(* IEC 61131-3 sources: volt/packages/volt-lsp-iec/test-corpus/lenze-mid/Device/Plc Logic/Application/A70_MachineModuleSources/MM_MachineControl/02_subMain, 11 files *)

(* ---- SidecorrectionCalculation.pou ---- *)
FUNCTION SidecorrectionCalculation
VAR_INPUT
	iAnalogInputValue						: INT;
	iSetpoint								: INT;
	iCorrectionScale						: REAL;
	iLightValue								: INT;
	iDarkValue								: INT;
	iNoWrapperOffsetPercentage01Perc		: INT; //test5

END_VAR
VAR_OUTPUT
	oIntPercentage							: INT;
	oRealPercentage							: REAL;
	oCorrectionValue						: REAL;
	oDeviationNoWrapper						: REAL;
END_VAR
VAR

	tRealMeasuredValue						: REAL;
	tRealPercentage							: REAL;
	tRealSetpoint							: REAL;
	tWhiteValue								: DINT;
	tBrownValue								: DINT;
	tWidthLight_Dark						: DINT;
	tRealWidthLight_Dark					: REAL;
	tMeasuredWithOffset						: REAL;
	tRealBrownValue							: REAL;
	tRealNoWrapperOffsetPercentage			: REAL;

END_VAR

%LANGUAGE ST
//Read out values for light and dark
tWhiteValue:=MOVE(iLightValue);
tBrownValue:=MOVE(iDarkValue);

//Calculate difference between light and dark value (light will be higher than dark)
tRealWidthLight_Dark:=TO_REAL(tWhiteValue-tBrownValue);
tRealBrownValue:=TO_REAL(tBrownValue);

//Measured value compensated with offset
tRealMeasuredValue:=TO_REAL(iAnalogInputValue);
tMeasuredWithOffset:=tRealMeasuredValue-tRealBrownValue;

//Calculation of the percentage
//"Measured value"/ Bandwidth
IF tRealWidthLight_Dark=0 THEN
	tRealWidthLight_Dark:=10;

END_IF
oRealPercentage:=(tMeasuredWithOffset/tRealWidthLight_Dark)*100;
oIntPercentage:=TO_INT(oRealPercentage);

//Calculation of the fault
//(act - set) * "correction scale"
tRealSetpoint:=TO_REAL(iSetpoint);
oCorrectionValue:=(oRealPercentage-tRealSetpoint)*iCorrectionScale;

//No wrapper detection
tRealNoWrapperOffsetPercentage:=TO_REAL(iNoWrapperOffsetPercentage01Perc);
oDeviationNoWrapper:=TO_INT(tRealNoWrapperOffsetPercentage*(tRealWidthLight_Dark/1000));

END_FUNCTION

(* ---- SpeedCalculationTrayfiller.pou ---- *)
FUNCTION SpeedCalculationTrayfiller
VAR_INPUT
END_VAR
VAR
	tInt: INT;
	tBool: BOOL;
END_VAR

%LANGUAGE LD
%NETWORK "NETWORK 1: Write setpoint speed in DB"
// The speed of the trayfiller has to be higher then the speed of the dryer. In this way there is always an empty space at the startpostition of the trayfiller.
MOVE(EN := ADD(EN := RAIL(), Mach1_Data.Drives.FeedForwardADS.Control.AutoSpeed, 30, OUT => tInt), tInt, OUT => Mach1_Data.Drives.FeedForwardATF.Control.AutoSpeed);
%NETWORK "NETWORK 2: Activation + Runtime guard feed forward dryer/trayfiller"
// Runtime calculation:
// 1 cycle = 60s/rpm
// speed = in 0.1 rpm -> 60s = 600 1/10s
//
// -> 1 cycle = 600/speed01
// DINT cannot calculate this 600/1000 = 0.1 -> DINT=0
// First multiply by 1000 (s -> ms)
// 1cycle = (600*1000)/speed1
// To give a little margin: add 500ms
ASSIGN(RuntimeGuard_V5_1_100(AlarmDB := Mach1_Alarms, iForward := Mach1_AuxData.TrayfillerActive AND Mach1_MIDS.IDB_TrayFiller.oFeedForwardMotor AND Mach1.Genflags.DelayAfterSTO AND (Mach1_AuxData.AllDrivesHomed OR INVERT(Mach1_AuxData.TrayfillerActive)), iReverse := LST_General.AlwaysOff, iActivateGuard := GE(EN := Mach1.Genflags.DelayAfterSTO AND Mach1_Data.Drives.FeedForwardATF.Control.StartAuto AND INVERT(LST_InputsOutputs.I133_3_PROX_zero_position_transport_ATF), Mach1_Data.Drives.FeedForwardATF.Control.AutoSpeed, 10).OUT, iMaxRuntime := T#10S, iReset := Mach1.GenFlags.StartFlag, iAlm := Mach1_Alarms.Alm051, ioAction := Mach1.GenFlags.MinorAlarm, ioAccRuntime := Mach1_AuxData.IEC_TIMERS.RuntimeGuardFeedforwardTrayfiller, oForwardGuarded => Mach1_Data.Drives.FeedForwardATF.Control.StartAuto), Q_SET => Mach1.GenFlags.StopDriveDirect);

END_FUNCTION

(* ---- Servo_LimitJog.pou ---- *)
FUNCTION_BLOCK Servo_LimitJog
VAR_INPUT
	iServoStatus 	: sUDT_ServoComm_Drive_Status;
	iServoControl 		: sUDT_ServoComm_Drive_Control;
END_VAR
VAR_OUTPUT
	oServoControl 		: sUDT_ServoComm_Drive_Control;
END_VAR
VAR
END_VAR
VAR_IN_OUT
	ioUDT_ServoDrive			: UDT_ServoDrive;
	ioUDT_JogLimitFree			: UDT_ServoJogLimitFree;
END_VAR

%LANGUAGE LD
%NETWORK "NETWORK 3 (p1): Check for limit switch"
ASSIGN(iServoStatus.Spare1, Q => ioUDT_JogLimitFree.Status.Limit_Left_OK);
%NETWORK "NETWORK 3 (p2): Check for limit switch"
ASSIGN(iServoStatus.Spare2, Q => ioUDT_JogLimitFree.Status.Limit_Right_OK);
%NETWORK "COPY previous control word to current controlword"
EXECUTE(EN := RAIL(), 'oServoControl:=iServoControl;');
%NETWORK "NETWORK 4 (p1): ControlToFreeLimitSwitches"
ASSIGN(ioUDT_JogLimitFree.Status.Limit_Left_OK AND ioUDT_JogLimitFree.Control.Jog_LimitToLeft, Q => oServoControl.Spare1);
%NETWORK "NETWORK 4 (p2): ControlToFreeLimitSwitches"
ASSIGN(ioUDT_JogLimitFree.Status.Limit_Right_OK AND ioUDT_JogLimitFree.Control.Jog_LimitToRight, Q => oServoControl.Spare2);

END_FUNCTION_BLOCK

(* ---- WSM.pou ---- *)
FUNCTION_BLOCK WSM
VAR_INPUT
	EN: BOOL;
	iGenflags : UDT_GeneralFlags;
	iInit: BOOL;
	iTest_Prod: BOOL;
	iCleaning: BOOL;
	iBunchPresent: BOOL;
	iWrapperPresentForLeafCarrier: BOOL;
	iPhotocellWrapper: BOOL;
	iWaterLevelSensor: BOOL;
	iTakeOverCycle: BOOL;
	iTimeOutSupplyWrapper: TIME;
	iSprayTime: TIME;
	iDelayContSpraying: TIME;
	iScreenForOperatorSettingsActivated: BOOL;
	iManualSprayCycleReset: BOOL;
	iManualSprayCycleStart: BOOL;
	iManualSprayCycleStop: BOOL;
	iMaxNumberOfSprayPulses: INT;

END_VAR
VAR_OUTPUT
	ENO: BOOL;
	oVentilationMotor: BOOL;
	oPositionMotor: BOOL;
	oWindingMotor: BOOL;
	oSprayingValve: BOOL;
	oWaterLevelValve: BOOL;
	oFaultWaitingForWrapper: BOOL;
	oFaultNoWrapper: BOOL;
	oFaultPhotocellWrapper : BOOL;
END_VAR
VAR
	stOSN_TakeOverCycle: F_TRIG;
	TMR_TimeOutSupply: TON;
	TMR_TimeOutPhotocell: TON;
	stRePositionMotor: R_TRIG;
	stSprayCycleActive: BOOL;
	TMR_DelayContinuousSpraying: TON;
	TMR_SprayTime: TON;
	stManualSprayCycleStarted: BOOL;

	TMR_ManualSprayCycleIdle: TON;

END_VAR

VAR_IN_OUT
	ioEnableSpraying: BOOL;
	ioManualSprayCycleActualCount: INT;
	ioManualStartSupply: BOOL;
END_VAR
VAR RETAIN PERSISTENT
	stRestposition: BOOL;
	stSupplyWrapper: BOOL;
	stWrapperPresent: BOOL;
	stNoWrapper: BOOL;
	stPhotocellWrapperFault: BOOL;
	stFeedForward: BOOL;
END_VAR
%LANGUAGE LD
%NETWORK "DONE Network 2: State: Initialise"
VAR w1 : ANY; END_VAR
w1 := iInit OR INVERT(iTest_Prod) OR iCleaning OR ioManualStartSupply;
ASSIGN(w1, Q_SET => stRestposition);
ASSIGN(w1, Q_RESET => stSupplyWrapper, Q_RESET => stWrapperPresent, Q_RESET => stNoWrapper, Q_RESET => stPhotocellWrapperFault);
%NETWORK "DONE Network 3: State: Restposition"
ASSIGN(stOSN_TakeOverCycle(CLK := iTakeOverCycle) AND stWrapperPresent, Q_SET => stRestposition, Q_RESET => stWrapperPresent);
%NETWORK "DONE Network 4: State: Supply wrapper"
ASSIGN(stRestposition AND (iTest_Prod AND INVERT(iCleaning) AND iBunchPresent AND INVERT(iTakeOverCycle) AND (iGenFlags.RunMan OR iGenFlags.RunAuto) OR ioManualStartSupply) OR stNoWrapper AND iGenFlags.StartFlag OR stPhotocellWrapperFault AND iGenFlags.StartFlag, Q_SET => stSupplyWrapper, Q_RESET => stRestposition, Q_RESET => stNoWrapper, Q_RESET => stPhotocellWrapperFault, Q_RESET => ioManualStartSupply);
%NETWORK "DONE Network 5: State: Wrapper Present"
VAR w2 : ANY; END_VAR
w2 := iWrapperPresentForLeafCarrier AND stSupplyWrapper;
ASSIGN(w2, Q_SET => stWrapperPresent);
ADD(EN := w2, 1, HMI_Var.Mach1.PRDWrapCurrentCntr, OUT => HMI_Var.Mach1.PRDWrapCurrentCntr);
ADD(EN := w2, 1, HMI_Var.Mach1.PRDWrapDayCounter, OUT => HMI_Var.Mach1.PRDWrapDayCounter);
ASSIGN(w2, Q_RESET => stSupplyWrapper);
%NETWORK "DONE Network 6: State: No Wrapper"
ASSIGN(TMR_TimeOutSupply(IN := stSupplyWrapper AND stFeedForward, PT := iTimeOutSupplyWrapper), Q_SET => stNoWrapper, Q_RESET => stSupplyWrapper);
%NETWORK "DONE Network 7: State: Photocell wrapper fault"
ASSIGN(TMR_TimeOutPhotocell(IN := stSupplyWrapper AND stFeedForward AND iPhotocellWrapper, PT := T#10S), Q_SET => stPhotocellWrapperFault, Q_RESET => stSupplyWrapper);
%NETWORK "DONE Network 8: Faults"
VAR w3 : ANY; END_VAR
w3 := True;
ASSIGN(w3 AND stSupplyWrapper AND iTakeOverCycle, Q => oFaultWaitingForWrapper);
ASSIGN(w3 AND stNoWrapper, Q => oFaultNoWrapper);
ASSIGN(w3 AND stPhotocellWrapperFault, Q => oFaultPhotocellWrapper);
%NETWORK "DONE Network 9: Ventilation motor"
ASSIGN(iGenFlags.EnableAuxDrive AND iTest_Prod AND INVERT(iCleaning), Q => oVentilationMotor);
%NETWORK "DONE Network 10:"
VAR w4 : ANY; END_VAR
w4 := iGenFlags.EnableAuxDrive AND stSupplyWrapper AND INVERT(iGenFlags.StopFlag);
ASSIGN(w4, Q => stFeedForward);
ASSIGN(w4, Q => oPositionMotor);
%NETWORK "DONE Network 11: Winding motor"
ASSIGN(iGenFlags.EnableAuxDrive AND INVERT(iGenFlags.StopFlag) AND iTest_Prod AND INVERT(iCleaning), Q => oWindingMotor);
%NETWORK "DONE Network 12: Start spray cycle"
VAR w5 : ANY; END_VAR
w5 := stFeedForward;
ASSIGN(stRePositionMotor(CLK := w5), Q_SET => stSprayCycleActive);
ASSIGN(TMR_DelayContinuousSpraying(IN := w5, PT := iDelayContSpraying), Q_SET => stSprayCycleActive);
%NETWORK "DONE Network 13: Timing spray cycle"
ASSIGN(TMR_SprayTime(IN := stSprayCycleActive, PT := iSprayTime) AND INVERT(TMR_DelayContinuousSpraying.Q), Q_RESET => stSprayCycleActive);
%NETWORK "DONE Network 14: Spraying valve"
ASSIGN(ioEnableSpraying AND stSprayCycleActive, Q => oSprayingValve);
%NETWORK "DONE Network 15: Automatic trigger of water"
ASSIGN(FALSE AND iGenFlags.EnablePneumEStop AND iWrapperPresentForLeafCarrier AND iTest_Prod AND INVERT(iCleaning), Q_SET => ioEnableSpraying);
%NETWORK "DONE Network 16: Water level control"
ASSIGN(ioEnableSpraying AND iWaterLevelSensor, Q => oWaterLevelValve);
%NETWORK "DONE Network 17: Manual spray cycle"
VAR w6 : ANY; END_VAR
w6 := iScreenForOperatorSettingsActivated;
MOVE(EN := w6 AND iManualSprayCycleReset, 0, OUT => ioManualSprayCycleActualCount);
ASSIGN(LT(EN := w6 AND iGenFlags.EnablePneumEStop AND (iManualSprayCycleStart OR stManualSprayCycleStarted) AND INVERT(iManualSprayCycleStop) AND INVERT(iManualSprayCycleReset), ioManualSprayCycleActualCount, iMaxNumberOfSprayPulses).OUT, Q => stManualSprayCycleStarted);
ASSIGN(ADD(EN := TMR_ManualSprayCycleIdle(IN := w6 AND stManualSprayCycleStarted AND INVERT(stSprayCycleActive), PT := T#300MS), ioManualSprayCycleActualCount, 1, OUT => ioManualSprayCycleActualCount), Q_SET => stSprayCycleActive);
%NETWORK "DONE Network 18: SAVE RLO"
ASSIGN(EN, Q => ENO);

END_FUNCTION_BLOCK

(* ---- AHWF.pou ---- *)
PROGRAM AHWF
VAR
	tFaultWaitingForWrapper : BOOL;
	tFaultNoWrapper: BOOL;
	tFaultPhotocellWrapper: BOOL;
	tStartFastWinding: BOOL;
	tSupplyWrapper: BOOL;
	tSprayingValve: BOOL;
	ttest: BOOL;
	R_TrigStartPos: R_TRIG;
END_VAR

VAR
	IDB_WSM: WSM;
END_VAR
%LANGUAGE LD
%NETWORK "Network 1: Detection of wrapper (set and reset)"
VAR w1 : ANY; END_VAR
w1 := True;
ASSIGN(w1 AND LST_InputsOutputs.I101_0_Wrapper_present, Q_SET => Mach1_AuxData.MemWrapperPassedUnderTheSensor);
ASSIGN(w1 AND INVERT(LST_InputsOutputs.I101_0_Wrapper_present) AND Mach1_AuxData.MemWrapperPassedUnderTheSensor, Q_SET => Mach1_AuxData.MemWrapperPresentForLeafCarrier, Q_SET => Mach1_AuxData.MemWrapperDetected_ResetLimitedSpeed);
ASSIGN(fc_CamC_CP_UDT(iEN := MOVE(EN := w1, Mach1_Data.CamControls.TakeOverCycle_C.Stop, OUT => Mach1_AuxData.CamControls.TakeOverCycleStopPulse_CP.Start), iMachinePosition := HMI_Var.Mach1.Position, iResetFlag := Mach1.GenFlags.Rotflag, ioPulse := Mach1_AuxData.CamControls.TakeOverCycleStopPulse_CP), Q_RESET => Mach1_AuxData.MemWrapperPresentForLeafCarrier, Q_RESET => Mach1_AuxData.MemWrapperPassedUnderTheSensor);
%NETWORK
ASSIGN(R_TrigStartPos(CLK := HMI_Var.HMI_AHWF_StartPos), Q_RESET => Mach1_AuxData.MemWrapperPresentForLeafCarrier, Q_RESET => Mach1_AuxData.MemWrapperPassedUnderTheSensor);
%NETWORK "Network 2: FB for DTA"
ASSIGN(IDB_WSM(EN := RAIL(), iGenflags := Mach1.GenFlags, iInit := LST_General.FirstCycle, iTest_Prod := HMI_Var.Test_Prod, iCleaning := HMI_Var.Btn_Cleaning, iBunchPresent := Mach1_AuxData.ShiftRegister.SR_bunch_present_position_1_JL, iWrapperPresentForLeafCarrier := Mach1_AuxData.MemWrapperPresentForLeafCarrier AND INVERT(HMI_Var.HMI_AHWF_fast_winding), iPhotocellWrapper := LST_InputsOutputs.I101_0_Wrapper_present AND INVERT(HMI_Var.HMI_AHWF_fast_winding), iWaterLevelSensor := LST_InputsOutputs.I101_3_Water_level_control, iTakeOverCycle := fc_CamC_CC_UDT(iEnable := True, iMachinePosition := HMI_Var.Mach1.Position, ioCamControl := Mach1_Data.CamControls.TakeOverCycle_C), iTimeOutSupplyWrapper := OPERAND('fc_dinttotime(Mach1_Data.Timers.TimeOutSupplyWrapper,2)'), iSprayTime := OPERAND('fc_dinttotime(Mach1_Data.Timers.SprayPulseWidth,2)'), iDelayContSpraying := OPERAND('fc_dinttotime(Mach1_Data.Timers.DelayContSpraying,2)'), iScreenForOperatorSettingsActivated := Mach1_AuxData.ScreenForOperatorSettingsActivated, iManualSprayCycleReset := HMI_Var.Mach1.SprayReset, iManualSprayCycleStart := HMI_Var.Mach1.SprayStart, iManualSprayCycleStop := HMI_Var.Mach1.SprayStop, iMaxNumberOfSprayPulses := Mach1_Data.Settings.Ints.MaxNumberOfSprayPulses, ioEnableSpraying := HMI_Var.Btn_Spraying, ioManualSprayCycleActualCount := Mach1_Data.Settings.Ints.ActualNumberOfSprayPulses, ioManualStartSupply := HMI_Var.HMI_AHWF_StartPos, oPositionMotor => tSupplyWrapper, oSprayingValve => tSprayingValve, oWaterLevelValve => LST_InputsOutputs.Q101_1_PNV_Waterlevel_control, oFaultWaitingForWrapper => tFaultWaitingForWrapper, oFaultNoWrapper => tFaultNoWrapper, oFaultPhotocellWrapper => tFaultPhotocellWrapper) AND Mach1.GenFlags.EnablePneumPressurised AND Mach1_Safety.Status.AllDoorsActuallyClosed AND tSprayingValve AND INVERT(Mach1_Alarms.Alm011), Q => PneumValveTerminalSMC.Pos1B);
%NETWORK "Network 3: Wrapper faults"
ASSIGN(Alarms_V5_1_100(AlarmDB := Mach1_Alarms, iCond := Mach1.GenFlags.DelayAfterEmergStop AND HMI_Var.Test_Prod AND INVERT(HMI_Var.Btn_Cleaning) AND tFaultWaitingForWrapper AND Mach1_AuxData.AllDrivesHomed, iReset := True, iAlm := Mach1_Alarms.Alm076, ioAction := Mach1.GenFlags.Warning) OR Alarms_V5_1_100(AlarmDB := Mach1_Alarms, iCond := Mach1.GenFlags.DelayAfterEmergStop AND HMI_Var.Test_Prod AND INVERT(HMI_Var.Btn_Cleaning) AND tFaultNoWrapper AND Mach1_AuxData.AllDrivesHomed, iReset := Mach1.GenFlags.StartFlag, iAlm := Mach1_Alarms.Alm043, ioAction := Mach1.GenFlags.MinorAlarm) OR Alarms_V5_1_100(AlarmDB := Mach1_Alarms, iCond := Mach1.GenFlags.DelayAfterEmergStop AND HMI_Var.Test_Prod AND INVERT(HMI_Var.Btn_Cleaning) AND INVERT(Mach1_Alarms.Alm045) AND tFaultPhotocellWrapper AND Mach1_AuxData.AllDrivesHomed, iReset := Mach1.GenFlags.StartFlag, iAlm := Mach1_Alarms.Alm045, ioAction := Mach1.GenFlags.MinorAlarm), Q_SET => Mach1.GenFlags.StopDriveDirect);
%NETWORK
%NETWORK "TODO Network 4: "
VAR w2 : ANY; w3 : ANY; w4 : ANY; END_VAR
w2 := True;
w3 := w2 AND True;
MOVE(EN := MOVE(EN := MOVE(EN := MOVE(EN := w3 AND TRUE, 175, OUT => Data_Exchange_Motion.FeedForwardWrapper.Control.VelUnit), 2000, OUT => Data_Exchange_Motion.FeedForwardWrapper.Control.DecUnit), 750, OUT => Data_Exchange_Motion.FeedForwardWrapper.Control.AccUnit), 100, OUT => Data_Exchange_Motion.FeedForwardWrapper.Control.TorqueLimit);
w4 := w3 AND HMI_Var.HMI_AHWF_fast_winding;
ASSIGN(Mach1_AuxData.IEC_TIMERS.TON_StartFastWinding(IN := w4, PT := T#200MS), Q => tStartFastWinding);
MOVE(EN := w4, 500, OUT => Data_Exchange_Motion.FeedForwardWrapper.Control.VelUnit);
MOVE(EN := w2, OPERAND('DINT_TO_LREAL(Mach1_Data.Settings.Dints.WrapperStopPosition)/10'), OUT => Data_Exchange_Motion.FeedForwardWrapper.Control.PosUnit);
ASSIGN(w2 AND INVERT(HMI_Var.HMI_AHWF_positioningType) AND INVERT(Mach1_Alarms.Alm056) AND mach1.Genflags.EnableAuxDrive AND (tSupplyWrapper OR tStartFastWinding OR Data_Exchange_Motion.FeedForwardWrapper.Control.StartTouchprobePos AND INVERT(Data_Exchange_Motion.FeedForwardWrapper.Status.InPosition)), Q => Data_Exchange_Motion.FeedForwardWrapper.Control.StartTouchprobePos);
ASSIGN(Mach1_AuxData.Edge.OSP_StopFlag(CLK := w2 AND (INVERT(Mach1_MIDS.FB_Mach1.iStop1) OR INVERT(Mach1_MIDS.FB_Mach1.iStop2) OR INVERT(Mach1_MIDS.FB_Mach1.iStop3) OR INVERT(Mach1_Safety.Status.AllDoorsActuallyClosed) OR LST_InputsOutputs.I101_0_Wrapper_present)), Q_RESET => HMI_Var.HMI_AHWF_fast_winding);
%NETWORK "Network 5: Side correction"
SideCorrection(EN := RAIL());
%NETWORK "Network 6: DTA-alarm: side limit reached"
ASSIGN(Alarms_V5_1_100(AlarmDB := Mach1_Alarms, iCond := Mach1_AuxData.Edge.OSP_LimitDTA_Reached(CLK := Mach1_AuxData.MIDS_Active AND Mach1.GenFlags.DelayAfterEmergStop AND (INVERT(Mach1_Data.Drives.SideCorrection_FreeLimit.Status.Limit_Left_OK) OR INVERT(Mach1_Data.Drives.SideCorrection_FreeLimit.Status.Limit_Right_OK))) AND Mach1_AuxData.AllDrivesHomed, iReset := Mach1.GenFlags.StartFlag, iAlm := Mach1_Alarms.Alm057, ioAction := Mach1.GenFlags.MinorAlarm) OR LST_General.AlwaysOff AND Alarms_V5_1_100(AlarmDB := Mach1_Alarms, iCond := Mach1_AuxData.MIDS_Active AND Mach1.GenFlags.DelayAfterEmergStop AND (INVERT(Mach1_Data.Drives.SideCorrection_FreeLimit.Status.Limit_Left_OK) OR INVERT(Mach1_Data.Drives.SideCorrection_FreeLimit.Status.Limit_Right_OK)) AND Mach1_AuxData.AllDrivesHomed, iReset := Mach1.GenFlags.StartFlag, iAlm := Mach1_Alarms.Alm074, ioAction := Mach1.GenFlags.Warning), Q_SET => Mach1.GenFlags.StopDriveDirect);
%NETWORK "Network 7: Alarm: Water receptacle full"
ASSIGN(Alarms_V5_1_100(AlarmDB := Mach1_Alarms, iCond := Mach1_AuxData.IEC_TIMERS.WaterReceptacleFull(IN := Mach1_AuxData.MIDS_Active AND LST_InputsOutputs.I101_3_Water_level_control AND INVERT(Mach1_Alarms.Alm055), PT := T#5M) AND HMI_Var.Test_Prod AND HMI_Var.Btn_Spraying AND Mach1_AuxData.AllDrivesHomed, iReset := Mach1.GenFlags.StartFlag, iAlm := Mach1_Alarms.Alm055, ioAction := Mach1.GenFlags.MinorAlarm), Q_SET => Mach1.GenFlags.StopDriveDirect);

END_PROGRAM

(* ---- fc_CheckRegister.pou ---- *)
PROGRAM fc_CheckRegister
VAR
END_VAR

%LANGUAGE LD
%NETWORK "NETWORK 1: Shift CheckRegister"
fc_ShiftRegister(ioPositie := db_CheckRegister.Positie);
%NETWORK "NETWORK 2: Check for error in dryer"
fc_CheckNumberOfErrorsRegister(iPositie := db_CheckRegister.Positie, iPositionToCheck := CTE.posCigarPresentOutfeed, iAmountOfErrors := Mach1_Data.Counters.MaxRepetitionNoCigarsDryer.SetValue, oError => db_CheckRegister.CheckRegisterError);

END_PROGRAM

(* ---- fc_Visualisation_HMI.pou ---- *)
PROGRAM fc_Visualisation_HMI
VAR_INPUT
END_VAR
VAR
	tbool: BOOL;
END_VAR

%LANGUAGE LD
%NETWORK "NETWORK 5: (P1) Visualisation - emergency stop"
Alarms_V5_1_100(AlarmDB := Mach1_Alarms, iCond := Mach1_AuxData.MIDS_Active AND INVERT(Mach1_Safety.Status.Emergency_button01), iReset := True, iAlm := Mach1_Alarms.Alm080, ioAction := Mach1.GenFlags.warning);
%NETWORK "NETWORK 5: (P2) Visualisation - emergency stop"
Alarms_V5_1_100(AlarmDB := Mach1_Alarms, iCond := Mach1_AuxData.MIDS_Active AND INVERT(Mach1_Safety.Status.Emergency_button02), iReset := True, iAlm := Mach1_Alarms.Alm081, ioAction := Mach1.GenFlags.warning);
%NETWORK "NETWORK 5: (P3) Visualisation - emergency stop"
Alarms_V5_1_100(AlarmDB := Mach1_Alarms, iCond := Mach1_AuxData.MIDS_Active AND INVERT(Mach1_Safety.Status.Emergency_button04), iReset := True, iAlm := Mach1_Alarms.Alm082, ioAction := Mach1.GenFlags.warning);
%NETWORK "DONE NETWORK 5 (p2): Visualisation - doors"
ASSIGN(Alarms_V5_1_100(AlarmDB := Mach1_Alarms, iCond := Mach1_AuxData.MIDS_Active AND Mach1.Genflags.DelayAfterEmergStop AND INVERT(Mach1_Safety.Status.Door_switch01), iReset := True, iAlm := Mach1_Alarms.Alm083, ioAction := Mach1.GenFlags.warning) OR Alarms_V5_1_100(AlarmDB := Mach1_Alarms, iCond := Mach1_AuxData.MIDS_Active AND Mach1.Genflags.DelayAfterEmergStop AND INVERT(Mach1_Safety.Status.Door_switch02), iReset := True, iAlm := Mach1_Alarms.Alm084, ioAction := Mach1.GenFlags.warning) OR Alarms_V5_1_100(AlarmDB := Mach1_Alarms, iCond := Mach1_AuxData.MIDS_Active AND Mach1.Genflags.DelayAfterEmergStop AND INVERT(Mach1_Safety.Status.Door_switch03), iReset := True, iAlm := Mach1_Alarms.Alm085, ioAction := Mach1.GenFlags.warning) OR Alarms_V5_1_100(AlarmDB := Mach1_Alarms, iCond := Mach1_AuxData.MIDS_Active AND Mach1.Genflags.DelayAfterEmergStop AND INVERT(Mach1_Safety.Status.Door_switch04), iReset := True, iAlm := Mach1_Alarms.Alm086, ioAction := Mach1.GenFlags.warning) OR Alarms_V5_1_100(AlarmDB := Mach1_Alarms, iCond := Mach1_AuxData.MIDS_Active AND Mach1.Genflags.DelayAfterEmergStop AND INVERT(Mach1_Safety.Status.Door_switch05), iReset := True, iAlm := Mach1_Alarms.Alm087, ioAction := Mach1.GenFlags.warning), Q => tbool);
%NETWORK
ASSIGN(Alarms_V5_1_100(AlarmDB := Mach1_Alarms, iCond := Mach1_AuxData.MIDS_Active AND Mach1.Genflags.DelayAfterEmergStop AND INVERT(Mach1_Safety.Status.Door_switch06), iReset := True, iAlm := Mach1_Alarms.Alm088, ioAction := Mach1.GenFlags.warning) OR Alarms_V5_1_100(AlarmDB := Mach1_Alarms, iCond := Mach1_AuxData.MIDS_Active AND Mach1.Genflags.DelayAfterEmergStop AND INVERT(Mach1_Safety.Status.Door_switch07), iReset := True, iAlm := Mach1_Alarms.Alm089, ioAction := Mach1.GenFlags.warning) OR Alarms_V5_1_100(AlarmDB := Mach1_Alarms, iCond := Mach1_AuxData.MIDS_Active AND Mach1.Genflags.DelayAfterEmergStop AND INVERT(Mach1_Safety.Status.Door_switch08), iReset := True, iAlm := Mach1_Alarms.Alm090, ioAction := Mach1.GenFlags.warning) OR Alarms_V5_1_100(AlarmDB := Mach1_Alarms, iCond := Mach1_AuxData.MIDS_Active AND Mach1.Genflags.DelayAfterEmergStop AND INVERT(Mach1_Safety.Status.Door_switch09), iReset := True, iAlm := Mach1_Alarms.Alm091, ioAction := Mach1.GenFlags.warning) OR Alarms_V5_1_100(AlarmDB := Mach1_Alarms, iCond := Mach1_AuxData.MIDS_Active AND Mach1.Genflags.DelayAfterEmergStop AND INVERT(Mach1_Safety.Status.Door_switch10), iReset := True, iAlm := Mach1_Alarms.Alm092, ioAction := Mach1.GenFlags.warning), Q => tbool);
%NETWORK
ASSIGN(Alarms_V5_1_100(AlarmDB := Mach1_Alarms, iCond := Mach1_AuxData.MIDS_Active AND Mach1.Genflags.DelayAfterEmergStop AND INVERT(Mach1_Safety.Status.Door_switch14), iReset := True, iAlm := Mach1_Alarms.Alm093, ioAction := Mach1.GenFlags.warning) OR Alarms_V5_1_100(AlarmDB := Mach1_Alarms, iCond := Mach1_AuxData.MIDS_Active AND Mach1.Genflags.DelayAfterEmergStop AND INVERT(Mach1_Safety.Status.Door_switch15), iReset := True, iAlm := Mach1_Alarms.Alm094, ioAction := Mach1.GenFlags.warning) OR Alarms_V5_1_100(AlarmDB := Mach1_Alarms, iCond := Mach1_AuxData.MIDS_Active AND Mach1.Genflags.DelayAfterEmergStop AND INVERT(Mach1_Safety.Status.Door_switch16), iReset := True, iAlm := Mach1_Alarms.Alm095, ioAction := Mach1.GenFlags.warning) OR Alarms_V5_1_100(AlarmDB := Mach1_Alarms, iCond := Mach1_AuxData.MIDS_Active AND Mach1.Genflags.DelayAfterEmergStop AND INVERT(Mach1_Safety.Status.Door_switch11), iReset := True, iAlm := Mach1_Alarms.Alm070, ioAction := Mach1.GenFlags.warning) OR Alarms_V5_1_100(AlarmDB := Mach1_Alarms, iCond := Mach1_AuxData.MIDS_Active AND Mach1.Genflags.DelayAfterEmergStop AND INVERT(Mach1_Safety.Status.Door_switch12), iReset := True, iAlm := Mach1_Alarms.Alm071, ioAction := Mach1.GenFlags.warning), Q => tbool);
%NETWORK
Alarms_V5_1_100(AlarmDB := Mach1_Alarms, iCond := Mach1_AuxData.MIDS_Active AND Mach1.Genflags.DelayAfterEmergStop AND INVERT(Mach1_Safety.Status.Door_switch13), iReset := True, iAlm := Mach1_Alarms.Alm072, ioAction := Mach1.GenFlags.warning);
%NETWORK
ASSIGN(Alarms_V5_1_100(AlarmDB := Mach1_Alarms, iCond := Mach1_AuxData.MIDS_Active AND Mach1.Genflags.DelayAfterEmergStop AND LST_InputsOutputs.I100_3_Selector_switch_auto_manual_OP0a, iReset := True, iAlm := Mach1_Alarms.Alm018, ioAction := Mach1.GenFlags.warning) OR Alarms_V5_1_100(AlarmDB := Mach1_Alarms, iCond := Mach1_AuxData.MIDS_Active AND Mach1.Genflags.DelayAfterEmergStop AND LST_InputsOutputs.I132_3_SW_Auto_Man, iReset := True, iAlm := Mach1_Alarms.Alm019, ioAction := Mach1.GenFlags.warning), Q => tbool);
%NETWORK "Reset of alarmlogging"
ASSIGN(Alarms_ResetAlarmLogging(EN := HMI_Var.ResetAlarmLogging, AlarmDB := Mach1_Alarms), Q_RESET => HMI_Var.ResetAlarmLogging);
%NETWORK "Adding product counters$R$L"
ASSIGN(ADD(EN := ADD(EN := ADD(EN := HMI_Var.Mach1.PRDCounterIncr, HMI_Var.Mach1.PRDTotalCounter, 1, OUT => HMI_Var.Mach1.PRDTotalCounter), HMI_Var.Mach1.PRDCigDayCounter, 1, OUT => HMI_Var.Mach1.PRDCigDayCounter), HMI_Var.Mach1.PRDCigCurrentCntr, 1, OUT => HMI_Var.Mach1.PRDCigCurrentCntr), Q_RESET => HMI_Var.Mach1.PRDCounterIncr);
%NETWORK "Reset Day Counter$R$L"
ASSIGN(MOVE(EN := MOVE(EN := HMI_Var.Mach1.PRDDayCounterReset_01, 0, OUT => HMI_Var.Mach1.PRDWrapDayCounter), 0, OUT => HMI_Var.Mach1.PRDCigDayCounter), Q_RESET => HMI_Var.Mach1.PRDDayCounterReset_01);
%NETWORK "Reset Current Counter$R$L"
ASSIGN(MOVE(EN := MOVE(EN := HMI_Var.Mach1.PRDDayCounterReset, 0, OUT => HMI_Var.Mach1.PRDWrapCurrentCntr), 0, OUT => HMI_Var.Mach1.PRDCigCurrentCntr), Q_RESET => HMI_Var.Mach1.PRDDayCounterReset);
%NETWORK
PRG_AlarmsToDWord(EN := TRUE);

END_PROGRAM

(* ---- MainDrive.pou ---- *)
PROGRAM MainDrive
VAR_INPUT
END_VAR
VAR
	tInt: INT;
	tMainDriveRun: BOOL;
	tMainDriveJog: BOOL;
END_VAR

VAR_OUTPUT
	oMainDriveRun: BOOL;
	oMainDriveJog: BOOL;
END_VAR
%LANGUAGE LD
%NETWORK "DONE NETWORK 1: Delay after doors closed"
ASSIGN(Mach1_AuxData.IEC_TIMERS.TON_DelayAfterDoorsClosed(IN := Mach1.GenFlags.DelayAfterEmergStop AND Mach1_Safety.Status.AllDoorsActuallyClosed AND Mach1_Safety.Status.DoorsOK, PT := T#150MS), Q => Mach1_AuxData.DelayAfterDoorsActuallyClosed);
%NETWORK "DONE NETWORK 2: Activating main drive"
VAR w1 : ANY; w2 : ANY; w3 : ANY; w4 : ANY; END_VAR
w1 := TRUE;
MOVE(EN := w1, 0, OUT => tInt);
ASSIGN(w1 AND INVERT(HMI_Var.Test_Prod), Q_RESET => Mach1_AuxData.MemLowerSpeedBecauseOfNoWrapper);
w2 := w1 AND Mach1.GenFlags.EnableMainDrive AND Mach1.GenFlags.ConditionsReadyForOperation AND INVERT(Mach1.GenFlags.StopDriveDirect) AND Mach1_AuxData.AllDrivesInLock;
w3 := w2 AND Mach1.GenFlags.RunAuto;
ASSIGN(w3, Q => tMainDriveRun, Q => oMainDriveRun, Q => Mach1_Safety.Control.RequestAutoSpeed);
MOVE(EN := BRANCH(FEED := w3, INVERT(Mach1_AuxData.MemLowerSpeedBecauseOfNoWrapper), LE(EN := Mach1_AuxData.MemLowerSpeedBecauseOfNoWrapper, Mach1_Data.AUTOSPEED, 40).OUT) AND INVERT(HMI_Var.Btn_Cleaning), Mach1_Data.AUTOSPEED, OUT => tInt);
MOVE(EN := GT(EN := w3 AND Mach1_AuxData.MemLowerSpeedBecauseOfNoWrapper, Mach1_Data.AUTOSPEED, 40).OUT AND INVERT(HMI_Var.Btn_Cleaning), 30, OUT => tInt);
MOVE(EN := w3 AND HMI_Var.Btn_Cleaning, 6, OUT => tInt);
w4 := w2 AND Mach1.GenFlags.RunMan;
ASSIGN(w4, Q => tMainDriveJog, Q => oMainDriveJog, Q => Mach1_Safety.Control.RequestManSpeed);
MOVE(EN := w4, Mach1_Data.MANUALSPEED, OUT => tInt);
RPM_To_DriveSpeed(iEN := w1, iRPM := tInt, oDriveSpeed => Mach1_Data.Drives.MainDrive_VM.Control.DriveMasterSpeed);
%NETWORK "DONE NETWORK 3 : DriveIsRunning flag"
VAR w5 : ANY; END_VAR
w5 := TRUE;
ASSIGN(w5, Q_RESET => Mach1.GenFlags.StopDriveDirect);
ASSIGN(w5 AND (tMainDriveRun OR tMainDriveJog), Q => Mach1.GenFlags.DriveIsRunning);
ASSIGN(Mach1_AuxData.IEC_TIMERS.TOFF_MainDriveAtProductionSpeed(IN := Mach1_AuxData.IEC_TIMERS.TON_MainDriveAtProductionSpeed(IN := w5 AND tMainDriveRun, PT := T#200MS), PT := T#60MS), Q => Mach1.GenFlags.DriveAtSpeed);
%NETWORK "DONE NETWORK 4: Alarm: Main drive blocked"
ASSIGN(Alarms_V5_1_100(AlarmDB := Mach1_Alarms, iCond := LT(EN := Mach1_AuxData.IEC_TIMERS.TON_MainDriveBlocked(IN := oMainDriveRun, PT := T#12S), HMI_Var.Mach1.ActualSpeed, 5).OUT, iReset := Mach1.GenFlags.StartFlag, iAlm := Mach1_Alarms.Alm040, ioAction := Mach1.GenFlags.MinorAlarm) AND Mach1_Alarms.Alm040, Q_SET => Mach1.GenFlags.StopDriveDirect);
%NETWORK "DONE NETWORK 5: Manual brakerelease"
%DISABLED
VAR w6 : ANY; END_VAR
w6 := TRUE;
ASSIGN(w6 AND Mach1_Alarms.Alm001 AND HMI_Var.ReleaseBrake, Q => LST_InputsOutputs.Q101_0_REL_release_brake);
ASSIGN(w6 AND (INVERT(Mach1_Alarms.Alm001) OR Mach1_Alarms.Alm001 AND INVERT(Mach1.GenFlags.StartFlag)), Q_RESET => HMI_Var.ReleaseBrake);

END_PROGRAM

(* ---- PRG_AlarmsToDWord.pou ---- *)
PROGRAM PRG_AlarmsToDWord
VAR
END_VAR

%LANGUAGE ST
dwErrorWord1.0:=Mach1_Alarms.Alm001;
dwErrorWord1.1:=Mach1_Alarms.Alm002;
dwErrorWord1.2:=Mach1_Alarms.Alm003;
dwErrorWord1.3:=Mach1_Alarms.Alm004;
dwErrorWord1.4:=Mach1_Alarms.Alm005;
dwErrorWord1.5:=Mach1_Alarms.Alm006;
dwErrorWord1.6:=Mach1_Alarms.Alm007;
dwErrorWord1.7:=Mach1_Alarms.Alm008;
dwErrorWord1.8:=Mach1_Alarms.Alm009;
dwErrorWord1.9:=Mach1_Alarms.Alm010;
dwErrorWord1.10:=Mach1_Alarms.Alm011;
dwErrorWord1.11:=Mach1_Alarms.Alm012;
dwErrorWord1.12:=Mach1_Alarms.Alm013;
dwErrorWord1.13:=Mach1_Alarms.Alm014;
dwErrorWord1.14:=Mach1_Alarms.Alm015;
dwErrorWord1.15:=Mach1_Alarms.Alm016;
dwErrorWord1.16:=Mach1_Alarms.Alm017;
dwErrorWord1.17:=Mach1_Alarms.Alm018;
dwErrorWord1.18:=Mach1_Alarms.Alm019;
dwErrorWord1.19:=Mach1_Alarms.Alm020;
dwErrorWord1.20:=Mach1_Alarms.Alm021;
dwErrorWord1.21:=Mach1_Alarms.Alm022;
dwErrorWord1.22:=Mach1_Alarms.Alm023;
dwErrorWord1.23:=Mach1_Alarms.Alm024;
dwErrorWord1.24:=Mach1_Alarms.Alm025;
dwErrorWord1.25:=Mach1_Alarms.Alm026;
dwErrorWord1.26:=Mach1_Alarms.Alm027;
dwErrorWord1.27:=Mach1_Alarms.Alm028;
dwErrorWord1.28:=Mach1_Alarms.Alm029;
dwErrorWord1.29:=Mach1_Alarms.Alm030;
dwErrorWord1.30:=Mach1_Alarms.Alm031;
dwErrorWord1.31:=Mach1_Alarms.Alm032;

dwErrorWord2.0:=Mach1_Alarms.Alm033;
dwErrorWord2.1:=Mach1_Alarms.Alm034;
dwErrorWord2.2:=Mach1_Alarms.Alm035;
dwErrorWord2.3:=Mach1_Alarms.Alm036;
dwErrorWord2.4:=Mach1_Alarms.Alm037;
dwErrorWord2.5:=Mach1_Alarms.Alm038;
dwErrorWord2.6:=Mach1_Alarms.Alm039;
dwErrorWord2.7:=Mach1_Alarms.Alm040;
dwErrorWord2.8:=Mach1_Alarms.Alm041;
dwErrorWord2.9:=Mach1_Alarms.Alm042;
dwErrorWord2.10:=Mach1_Alarms.Alm043;
dwErrorWord2.11:=Mach1_Alarms.Alm044;
dwErrorWord2.12:=Mach1_Alarms.Alm045;
dwErrorWord2.13:=Mach1_Alarms.Alm046;
dwErrorWord2.14:=Mach1_Alarms.Alm047;
dwErrorWord2.15:=Mach1_Alarms.Alm048;
dwErrorWord2.16:=Mach1_Alarms.Alm049;
dwErrorWord2.17:=Mach1_Alarms.Alm050;
dwErrorWord2.18:=Mach1_Alarms.Alm051;
dwErrorWord2.19:=Mach1_Alarms.Alm052;
dwErrorWord2.20:=Mach1_Alarms.Alm053;
dwErrorWord2.21:=Mach1_Alarms.Alm054;
dwErrorWord2.22:=Mach1_Alarms.Alm055;
dwErrorWord2.23:=Mach1_Alarms.Alm056;
dwErrorWord2.24:=Mach1_Alarms.Alm057;
dwErrorWord2.25:=Mach1_Alarms.Alm058;
dwErrorWord2.26:=Mach1_Alarms.Alm059;
dwErrorWord2.27:=Mach1_Alarms.Alm060;
dwErrorWord2.28:=Mach1_Alarms.Alm061;
dwErrorWord2.29:=Mach1_Alarms.Alm062;
dwErrorWord2.30:=Mach1_Alarms.Alm063;
dwErrorWord2.31:=Mach1_Alarms.Alm064;

dwErrorWord3.0:=Mach1_Alarms.Alm065;
dwErrorWord3.1:=Mach1_Alarms.Alm066;
dwErrorWord3.2:=Mach1_Alarms.Alm067;
dwErrorWord3.3:=Mach1_Alarms.Alm068;
dwErrorWord3.4:=Mach1_Alarms.Alm069;
dwErrorWord3.5:=Mach1_Alarms.Alm070;
dwErrorWord3.6:=Mach1_Alarms.Alm071;
dwErrorWord3.7:=Mach1_Alarms.Alm072;
dwErrorWord3.8:=Mach1_Alarms.Alm073;
dwErrorWord3.9:=Mach1_Alarms.Alm074;
dwErrorWord3.10:=Mach1_Alarms.Alm075;
dwErrorWord3.11:=Mach1_Alarms.Alm076;
dwErrorWord3.12:=Mach1_Alarms.Alm077;
dwErrorWord3.13:=Mach1_Alarms.Alm078;
dwErrorWord3.14:=Mach1_Alarms.Alm079;
dwErrorWord3.15:=Mach1_Alarms.Alm080;
dwErrorWord3.16:=Mach1_Alarms.Alm081;
dwErrorWord3.17:=Mach1_Alarms.Alm082;
dwErrorWord3.18:=Mach1_Alarms.Alm083;
dwErrorWord3.19:=Mach1_Alarms.Alm084;
dwErrorWord3.20:=Mach1_Alarms.Alm085;
dwErrorWord3.21:=Mach1_Alarms.Alm086;
dwErrorWord3.22:=Mach1_Alarms.Alm087;
dwErrorWord3.23:=Mach1_Alarms.Alm088;
dwErrorWord3.24:=Mach1_Alarms.Alm089;
dwErrorWord3.25:=Mach1_Alarms.Alm090;
dwErrorWord3.26:=Mach1_Alarms.Alm091;
dwErrorWord3.27:=Mach1_Alarms.Alm092;
dwErrorWord3.28:=Mach1_Alarms.Alm093;
dwErrorWord3.29:=Mach1_Alarms.Alm094;
dwErrorWord3.30:=Mach1_Alarms.Alm095;
dwErrorWord3.31:=Mach1_Alarms.Alm096;

dwErrorWord4.0:=Mach1_Alarms.Alm097;
dwErrorWord4.1:=Mach1_Alarms.Alm098;
dwErrorWord4.2:=Mach1_Alarms.Alm099;
dwErrorWord4.3:=Mach1_Alarms.Alm100;

END_PROGRAM

(* ---- SideCorrection.pou ---- *)
PROGRAM SideCorrection
VAR_INPUT
END_VAR
VAR
	tCorrectionScale			: DINT;
	tCorrectionScaleReal		: REAL;
	tReal						: REAL;
	tDint						: DINT;
	tInt						: INT;

	tbool: BOOL;
END_VAR

%LANGUAGE LD
%NETWORK "Network 1: Averaging of sensorsignal"
fc_MeanValue(EN := RAIL(), iLength := 20, iAcquireNewValue := True, iNewValue := OPERAND('TO_INT(LST_InputsOutputs.IW340_LeafCoverageSensor)'), ioValues := db_MeanValuesSideCorrectionSensor.MeasurementValues, oMeanValue => DB_Kantcorrectie.MeasuredValue);
%NETWORK
VAR w1 : ANY; END_VAR
w1 := TRUE;
ASSIGN(MOVE(EN := w1 AND DB_Kantcorrectie.CopyMeasuredToDark, DB_Kantcorrectie.MeasuredValue, OUT => DB_Kantcorrectie.DarkValue), Q_RESET => DB_Kantcorrectie.CopyMeasuredToDark);
ASSIGN(MOVE(EN := w1 AND DB_Kantcorrectie.CopyMeasuredToLight, DB_Kantcorrectie.MeasuredValue, OUT => DB_Kantcorrectie.LightValue), Q_RESET => DB_Kantcorrectie.CopyMeasuredToLight);
%NETWORK "Network 2: Read out inputvalue and calculate correctionvalue"
MOVE(EN := SidecorrectionCalculation(EN := MOVE(EN := TRUE, Mach1_Data.Settings.Ints.SideCorrectionScaleFactor, OUT => tCorrectionScale), iAnalogInputValue := DB_Kantcorrectie.MeasuredValue, iSetpoint := DB_Kantcorrectie.Setpoint, iCorrectionScale := -1, iLightValue := DB_Kantcorrectie.LightValue, iDarkValue := DB_Kantcorrectie.DarkValue, iNoWrapperOffsetPercentage01Perc := DB_Kantcorrectie.NoWrapperPercentage, oIntPercentage => DB_Kantcorrectie.Percentage10, oCorrectionValue => DB_Kantcorrectie.MeasuredValueReal, oDeviationNoWrapper => tReal), OPERAND('REAL_TO_INT(tReal)'), OUT => DB_Kantcorrectie.DeviationNoWrapper);
%NETWORK "Network 3: Determine side-correction value"
VAR w2 : ANY; w3 : ANY; END_VAR
w2 := fc_CamC_CP_UDT(iEN := RAIL(), iMachinePosition := HMI_Var.Mach1.Position, iResetFlag := Mach1.GenFlags.Rotflag, ioPulse := Mach1_Data.CamControls.MeasurementForSidecorrection_CP);
MOVE(EN := MOVE(EN := w2 AND Mach1_Data.Drives.SideCorrection_FreeLimit.Status.Limit_Left_OK AND Mach1_Data.Drives.SideCorrection_FreeLimit.Status.Limit_right_OK, DB_Kantcorrectie.MeasuredValueReal, OUT => DB_Kantcorrectie.CopiedValueReal), DB_Kantcorrectie.Percentage10, OUT => DB_Kantcorrectie.CopiedValueInt);
w3 := w2 AND Mach1_AuxData.MemWrapperDetected_ResetLimitedSpeed;
ASSIGN(w3, Q_RESET => Mach1_AuxData.MemLowerSpeedBecauseOfNoWrapper);
ASSIGN(w3, Q_RESET => Mach1_AuxData.MemWrapperDetected_ResetLimitedSpeed);
ASSIGN(GT(EN := SUB(EN := w2, DB_Kantcorrectie.LightValue, DB_Kantcorrectie.DeviationNoWrapper, OUT => DB_Kantcorrectie.NoWrapperValue), LST_InputsOutputs.IW340_LeafCoverageSensor, DB_Kantcorrectie.NoWrapperValue).OUT AND HMI_Var.Test_Prod, Q_SET => Mach1_AuxData.MemLowerSpeedBecauseOfNoWrapper);
%NETWORK "DONE Network 4: In case a limit switch is reached: overwrite values"
VAR w4 : ANY; END_VAR
w4 := True;
MOVE(EN := w4 AND INVERT(Mach1_Data.Drives.SideCorrection_FreeLimit.Status.Limit_Left_OK) AND Mach1_Data.Drives.SideCorrection_FreeLimit.Status.Limit_Right_OK, -100.0, OUT => DB_Kantcorrectie.CopiedValueReal);
MOVE(EN := MOVE(EN := w4 AND INVERT(Mach1_Data.Drives.SideCorrection_FreeLimit.Status.Limit_Right_OK) AND Mach1_Data.Drives.SideCorrection_FreeLimit.Status.Limit_Left_OK, 100.0, OUT => DB_Kantcorrectie.CopiedValueReal), -1, OUT => tCorrectionScale);
MOVE(EN := MOVE(EN := w4 AND (INVERT(Mach1_Data.Drives.SideCorrection_FreeLimit.Status.Limit_Left_OK) AND INVERT(Mach1_Data.Drives.SideCorrection_FreeLimit.Status.Limit_Right_OK) OR INVERT(HMI_Var.Test_Prod) OR Mach1_AuxData.MemLowerSpeedBecauseOfNoWrapper), 0.0, OUT => DB_Kantcorrectie.CopiedValueReal), 1, OUT => tCorrectionScale);
%NETWORK "DONE Network 5: Write side-correction values to the servo drive"
EXECUTE(EN := RAIL(), 'tReal:=DB_Kantcorrectie.CopiedValueReal*DINT_TO_REAL(tCorrectionScale);
Mach1_Data.Drives.SideCorrection.CAM.Y_Scale_Recipe:=REAL_TO_INT(tReal/(-1000));
');
%NETWORK "DONE Network 6 : Manual adjustment of the sidecorrection"
VAR w5 : ANY; END_VAR
w5 := True;
ASSIGN(w5 AND Mach1_Data.Drives.SideCorrection_FreeLimit.Status.Limit_Left_OK AND HMI_Var.Mach1.DTA_PositioningLeft, Q => Mach1_Data.Drives.SideCorrection_FreeLimit.Control.Jog_LimitToLeft);
ASSIGN(w5 AND Mach1_Data.Drives.SideCorrection_FreeLimit.Status.Limit_Right_OK AND HMI_Var.Mach1.DTA_PositioningRight, Q => Mach1_Data.Drives.SideCorrection_FreeLimit.Control.Jog_LimitToRight);

END_PROGRAM

(* ---- SpeedCalculationDryer.pou ---- *)
PROGRAM SpeedCalculationDryer
VAR_INPUT
END_VAR
VAR
	TempI: INT;
	cor_DenumI: INT:=1;
	cor_NumI: INT:=1;
	cor_DenumDI: DINT:=1;
	cor_NumDI: DINT:=1;
	Speed01rpm: INT;
	tSetHighSpeedCycles : BOOL;
	cor_Const: INT;
	R_TRIG_0: R_TRIG;
	MainDrive_AutoSpeed01rpm: INT;
	Mach_ActSpeed_Rpm01:INT;
	devAngle: INT;

END_VAR

%LANGUAGE LD
%NETWORK "NETWORK 1 : Speed control transport system dryer"
VAR w1 : ANY; w2 : ANY; w3 : ANY; w4 : ANY; END_VAR
w1 := True;
MOVE(EN := w1, 0, OUT => TempI);
MUL(EN := w1, Mach1_Data.AUTOSPEED, 10, OUT => MainDrive_AutoSpeed01rpm);
MOVE(EN := w1, MainDrive_AutoSpeed01rpm, OUT => Droger_Data.Cor_denumerator);
w2 := w1 AND True;
MOVE(EN := MOVE(EN := Mach1_AuxData.IEC_TIMERS.TON_DelayIdling(IN := w2 AND INVERT(Mach1.GenFlags.DriveIsRunning), PT := T#500MS) AND INVERT(Mach1_Alarms.Alm049), MainDrive_AutoSpeed01rpm, OUT => Mach_ActSpeed_Rpm01), MainDrive_AutoSpeed01rpm, OUT => Droger_Data.Cor_numerator);
MOVE(EN := w2 AND (Mach1.GenFlags.DriveIsRunning OR INVERT(Mach1_AuxData.IEC_TIMERS.TON_DelayIdling.Q)), OPERAND('HMI_Var.Mach1.ActualSpeed*10'), OUT => Mach_ActSpeed_Rpm01);
w3 := w2 AND True;
w4 := w3 AND Trayfiller_Data.commInterface.HoldFeedFwd;
MOVE(EN := ASSIGN(w4 AND (LST_InputsOutputs.I133_1_PROX_zero_position_transport_ADS OR Mach1_AuxData.ADS_StopOnZeroPulse), Q => Mach1_AuxData.ADS_StopOnZeroPulse), 750, OUT => Droger_Data.Cor_numerator);
MOVE(EN := Mach1_AuxData.Edge.Osr_SetCounter(CLK := w4 AND Trayfiller_Data.commInterface.Permission), 5, OUT => Mach1_AuxData.CounterHighSpeedATF_ADS);
MUL(EN := NE(EN := w3 AND Trayfiller_Data.commInterface.Permission, Mach1_AuxData.CounterHighSpeedATF_ADS, 0).OUT, Mach1_Data.AUTOSPEED, 13, OUT => Droger_Data.Cor_numerator);
EXECUTE(EN := w2, 'cor_NumDI:=Droger_Data.Cor_numerator;
cor_DenumDI:=Droger_Data.Cor_denumerator;
//cor_NumDI:=1;
//cor_DenumDI:=1;
HMI_Var.Mach1.ActualSpeedDryer:=(Mach_ActSpeed_Rpm01*cor_numDI)/cor_denumdi;
Mach1_Data.Drives.FeedForwardADS.Control.AutoSpeed:=REAL_TO_INT(0.9*dint_to_real(HMI_Var.Mach1.ActualSpeedDryer)*6/10);

');
%NETWORK "NETWORK 2: Deviation calculation of sync point, transport system trayfiller"
VAR w5 : ANY; END_VAR
// Principle: It's better to accelerate the drive then to decelerate, because otherwise cigars could be missed.
// So that is why the deceleration should be kept short, by trial and error the optimum point is 60degrees (difference between setpoint and actual point).
// dev: [0-60]: dec.
// dev: ]60-360]: acc.
//
// Numerator = (Act_syncpos -/- Gew_syncpos) + Cte
// Cte=little bit slower then the value for the set speed. (If the mid-s rotates 100rpm (value=1000), then this value should be a little less (e.g 99,8rpm).
//         This way, the system lags a little bit, and therefor needs to accelerate (which is beter). If the system leads, then it needs to decel. (which is not ideal)
//
// Uit metingen is gebleken dat de optimale synchronisatiepositie op 60 graden
// ligt.
//
// correctie  -60     0     60     120    180    240    300
//             |------|------|------|------|------|------|--
// encoder     0     60     120    180    240    300    360
//
// Om de ingestelde synchronisatiepositie te verschuiven naar het optimale window
// van -60..300 wordt de correctiefactor gecorrigeerd:
//  - indien correctie < -60 dan 360 erbij optellen
//  - indien correctie > 300 dan 360 eraf tellen
w5 := ADD(EN := SUB(EN := SUB(EN := Mach1.GenFlags.DriveIsRunning, Droger_Data.Act_sync_pos, Droger_Data.set_sync_pos, OUT => devAngle), MainDrive_AutoSpeed01rpm, 2, OUT => cor_Const), devAngle, cor_Const, OUT => Droger_Data.Cor_numerator);
ADD(EN := LT(EN := w5, devAngle, -60).OUT, Droger_Data.Cor_numerator, 360, OUT => Droger_Data.Cor_numerator);
SUB(EN := GT(EN := w5, devAngle, 300).OUT, Droger_Data.Cor_numerator, 360, OUT => Droger_Data.Cor_numerator);
%NETWORK
VAR w6 : ANY; END_VAR
w6 := R_TRIG_0(CLK := LST_InputsOutputs.I133_1_PROX_zero_position_transport_ADS);
MOVE(EN := w6, HMI_Var.Mach1.Position, OUT => Droger_Data.Act_sync_pos);
MOVE(EN := w6, Mach1_Data.CamControls.FeedforwardDryer_CP.Start, OUT => Droger_Data.set_sync_pos);
SUB(EN := GT(EN := w6, Mach1_AuxData.CounterHighSpeedATF_ADS, 0).OUT, Mach1_AuxData.CounterHighSpeedATF_ADS, 1, OUT => Mach1_AuxData.CounterHighSpeedATF_ADS);

END_PROGRAM
